(* IEC 61131-3 sources: llm-plc-st-eval/codesys/dobles/A5, 9 files *)

(* ---- 01_Correcta.st ---- *)
(* DOBLE DE PRUEBA A5/Correcta - NO ES CORPUS. Esperado: veredicto 1 *)
TYPE ST_Evento :
STRUCT
    codigo : INT;
    marca : TIME;
END_STRUCT
END_TYPE

FUNCTION_BLOCK FB_Registro
VAR_INPUT
    evento : INT;
    nuevoEvento : BOOL;
    ciclo : TIME;
END_VAR
VAR_OUTPUT
    buffer : ARRAY[0..19] OF ST_Evento;
    indice : INT := -1;
    nEventos : INT;
END_VAR
VAR
    tAcum : TIME;
    prev : BOOL;
    nTotal : INT;
END_VAR
tAcum := tAcum + ciclo;
IF (nuevoEvento AND NOT prev) AND (TRUE) THEN
    indice := (indice + 1) MOD 20;
    buffer[indice].codigo := evento;
    buffer[indice].marca := tAcum;
    nEventos := MIN(20, nEventos + 1);
END_IF
prev := nuevoEvento;
END_FUNCTION_BLOCK

(* ---- 02_CorrectaAcumDespues.st ---- *)
(* DOBLE DE PRUEBA A5/CorrectaAcumDespues - NO ES CORPUS. Esperado: veredicto 1 *)
TYPE ST_Evento :
STRUCT
    codigo : INT;
    marca : TIME;
END_STRUCT
END_TYPE

FUNCTION_BLOCK FB_Registro
VAR_INPUT
    evento : INT;
    nuevoEvento : BOOL;
    ciclo : TIME;
END_VAR
VAR_OUTPUT
    buffer : ARRAY[0..19] OF ST_Evento;
    indice : INT := -1;
    nEventos : INT;
END_VAR
VAR
    tAcum : TIME;
    prev : BOOL;
    nTotal : INT;
END_VAR
IF (nuevoEvento AND NOT prev) AND (TRUE) THEN
    indice := (indice + 1) MOD 20;
    buffer[indice].codigo := evento;
    buffer[indice].marca := tAcum;
    nEventos := MIN(20, nEventos + 1);
END_IF
prev := nuevoEvento;
tAcum := tAcum + ciclo;
END_FUNCTION_BLOCK

(* ---- 03_IndiceInicialCero.st ---- *)
(* DOBLE DE PRUEBA A5/IndiceInicialCero - NO ES CORPUS. Esperado: veredicto 2, falla en el paso 0 *)
TYPE ST_Evento :
STRUCT
    codigo : INT;
    marca : TIME;
END_STRUCT
END_TYPE

FUNCTION_BLOCK FB_Registro
VAR_INPUT
    evento : INT;
    nuevoEvento : BOOL;
    ciclo : TIME;
END_VAR
VAR_OUTPUT
    buffer : ARRAY[0..19] OF ST_Evento;
    indice : INT;
    nEventos : INT;
END_VAR
VAR
    tAcum : TIME;
    prev : BOOL;
    nTotal : INT;
    vacio : BOOL := TRUE;
END_VAR
tAcum := tAcum + ciclo;
IF (nuevoEvento AND NOT prev) AND (TRUE) THEN
    indice := SEL(vacio, (indice + 1) MOD 20, 0);
    buffer[indice].codigo := evento;
    buffer[indice].marca := tAcum;
    nEventos := MIN(20, nEventos + 1);
    vacio := FALSE;
END_IF
prev := nuevoEvento;
END_FUNCTION_BLOCK

(* ---- 04_CuentaPorNivel.st ---- *)
(* DOBLE DE PRUEBA A5/CuentaPorNivel - NO ES CORPUS. Esperado: veredicto 2, falla en el paso 1 *)
TYPE ST_Evento :
STRUCT
    codigo : INT;
    marca : TIME;
END_STRUCT
END_TYPE

FUNCTION_BLOCK FB_Registro
VAR_INPUT
    evento : INT;
    nuevoEvento : BOOL;
    ciclo : TIME;
END_VAR
VAR_OUTPUT
    buffer : ARRAY[0..19] OF ST_Evento;
    indice : INT := -1;
    nEventos : INT;
END_VAR
VAR
    tAcum : TIME;
    prev : BOOL;
    nTotal : INT;
END_VAR
tAcum := tAcum + ciclo;
IF (nuevoEvento) AND (TRUE) THEN
    indice := (indice + 1) MOD 20;
    buffer[indice].codigo := evento;
    buffer[indice].marca := tAcum;
    nEventos := MIN(20, nEventos + 1);
END_IF
prev := nuevoEvento;
END_FUNCTION_BLOCK

(* ---- 05_MarcaSinAcumular.st ---- *)
(* DOBLE DE PRUEBA A5/MarcaSinAcumular - NO ES CORPUS. Esperado: veredicto 2, falla en el paso 1 *)
TYPE ST_Evento :
STRUCT
    codigo : INT;
    marca : TIME;
END_STRUCT
END_TYPE

FUNCTION_BLOCK FB_Registro
VAR_INPUT
    evento : INT;
    nuevoEvento : BOOL;
    ciclo : TIME;
END_VAR
VAR_OUTPUT
    buffer : ARRAY[0..19] OF ST_Evento;
    indice : INT := -1;
    nEventos : INT;
END_VAR
VAR
    tAcum : TIME;
    prev : BOOL;
    nTotal : INT;
END_VAR
tAcum := tAcum + ciclo;
IF (nuevoEvento AND NOT prev) AND (TRUE) THEN
    indice := (indice + 1) MOD 20;
    buffer[indice].codigo := evento;
    buffer[indice].marca := ciclo;
    nEventos := MIN(20, nEventos + 1);
END_IF
prev := nuevoEvento;
END_FUNCTION_BLOCK

(* ---- 06_PrimeroEnPosicion1.st ---- *)
(* DOBLE DE PRUEBA A5/PrimeroEnPosicion1 - NO ES CORPUS. Esperado: veredicto 2, falla en el paso 0 *)
TYPE ST_Evento :
STRUCT
    codigo : INT;
    marca : TIME;
END_STRUCT
END_TYPE

FUNCTION_BLOCK FB_Registro
VAR_INPUT
    evento : INT;
    nuevoEvento : BOOL;
    ciclo : TIME;
END_VAR
VAR_OUTPUT
    buffer : ARRAY[0..19] OF ST_Evento;
    indice : INT;
    nEventos : INT;
END_VAR
VAR
    tAcum : TIME;
    prev : BOOL;
    nTotal : INT;
END_VAR
tAcum := tAcum + ciclo;
IF (nuevoEvento AND NOT prev) AND (TRUE) THEN
    indice := (indice + 1) MOD 20;
    buffer[indice].codigo := evento;
    buffer[indice].marca := tAcum;
    nEventos := MIN(20, nEventos + 1);
END_IF
prev := nuevoEvento;
END_FUNCTION_BLOCK

(* ---- 07_SinSobrescritura.st ---- *)
(* DOBLE DE PRUEBA A5/SinSobrescritura - NO ES CORPUS. Esperado: veredicto 2, falla en el paso 4 *)
TYPE ST_Evento :
STRUCT
    codigo : INT;
    marca : TIME;
END_STRUCT
END_TYPE

FUNCTION_BLOCK FB_Registro
VAR_INPUT
    evento : INT;
    nuevoEvento : BOOL;
    ciclo : TIME;
END_VAR
VAR_OUTPUT
    buffer : ARRAY[0..19] OF ST_Evento;
    indice : INT := -1;
    nEventos : INT;
END_VAR
VAR
    tAcum : TIME;
    prev : BOOL;
    nTotal : INT;
END_VAR
tAcum := tAcum + ciclo;
IF (nuevoEvento AND NOT prev) AND (nEventos < 20) THEN
    indice := (indice + 1) MOD 20;
    buffer[indice].codigo := evento;
    buffer[indice].marca := tAcum;
    nEventos := MIN(20, nEventos + 1);
END_IF
prev := nuevoEvento;
END_FUNCTION_BLOCK

(* ---- 08_NEventosSinTope.st ---- *)
(* DOBLE DE PRUEBA A5/NEventosSinTope - NO ES CORPUS. Esperado: veredicto 2, falla en el paso 4 *)
TYPE ST_Evento :
STRUCT
    codigo : INT;
    marca : TIME;
END_STRUCT
END_TYPE

FUNCTION_BLOCK FB_Registro
VAR_INPUT
    evento : INT;
    nuevoEvento : BOOL;
    ciclo : TIME;
END_VAR
VAR_OUTPUT
    buffer : ARRAY[0..19] OF ST_Evento;
    indice : INT := -1;
    nEventos : INT;
END_VAR
VAR
    tAcum : TIME;
    prev : BOOL;
    nTotal : INT;
END_VAR
tAcum := tAcum + ciclo;
IF (nuevoEvento AND NOT prev) AND (TRUE) THEN
    indice := (indice + 1) MOD 20;
    buffer[indice].codigo := evento;
    buffer[indice].marca := tAcum;
    nEventos := nEventos + 1;
END_IF
prev := nuevoEvento;
END_FUNCTION_BLOCK

(* ---- 09_VueltaAPosicion1.st ---- *)
(* DOBLE DE PRUEBA A5/VueltaAPosicion1 - NO ES CORPUS. Esperado: veredicto 2, falla en el paso 4 *)
TYPE ST_Evento :
STRUCT
    codigo : INT;
    marca : TIME;
END_STRUCT
END_TYPE

FUNCTION_BLOCK FB_Registro
VAR_INPUT
    evento : INT;
    nuevoEvento : BOOL;
    ciclo : TIME;
END_VAR
VAR_OUTPUT
    buffer : ARRAY[0..19] OF ST_Evento;
    indice : INT := -1;
    nEventos : INT;
END_VAR
VAR
    tAcum : TIME;
    prev : BOOL;
    nTotal : INT;
END_VAR
tAcum := tAcum + ciclo;
IF (nuevoEvento AND NOT prev) AND (TRUE) THEN
    indice := SEL(indice < 19, 1, indice + 1);
    buffer[indice].codigo := evento;
    buffer[indice].marca := tAcum;
    nEventos := MIN(20, nEventos + 1);
END_IF
prev := nuevoEvento;
END_FUNCTION_BLOCK
